// Vereinfachter Achszustand für die GUI.
{attribute 'qualified_only'}
{attribute 'strict'}
{attribute 'to_string'}
TYPE E_AxisState :
(
    Disabled := 0,
    Standstill := 1,
    Moving := 2, // Einzelbewegung
    Coupled := 3, // über FB_BendKinematics gekoppelt
    Error := 4
) INT;
END_TYPE

(* stored: Version 1.1.0.1
   DUT E_AxisState: Id {ce9c02e4-aafb-4062-97ff-bbaaeca05990} *)
